(* IEC 61131-3 sources: codesys-to-s7/tests/corpus/C2S7-TYPE-RANGE/neg, 1 file *)

(* ---- input.st ---- *)
FUNCTION_BLOCK FB_Case
VAR
    x : INT;
END_VAR
x := 5;
END_FUNCTION_BLOCK
